// SIMATIC S7-200 project (STEP 7-Micro/WIN), CPU 224 CN REL 02.01

SYMBOL_TABLE USUARIO1
SM2              I0.0     // Sensor magnetico extendido del cilindro retenedor
SM1              I0.1     // Sensor magnetico retraido del cilindor retenedor
SM4              I0.2     // Sensor magnetico extendido del cilindro de empuje
SM3              I0.3     // Sensor magnetico retraido del cilindor de empuje
SF               I0.4     // Sensor Fotoelectrico Final
SP               I0.5     // Sensor Fotoelectrico Superior
SP1              I0.6     // Sensor Fotoelectrico Inferior
SII              I0.7     // Sensor Inductivo
SB_1             I1.2     // Pulsador de marcha
SB_2             I1.3     // Pulsador de paro
QS               I1.4     // Zeta de Emergencia
SA               I1.5     // Selector de modo
KV1              Q0.0     // Cilindro neumatico Retenedor
KV2              Q0.1     // Cilindro neumatico de empuje
HL1              Q0.7     // Señalizacion amarillo
HL2              Q1.0     // Señalizacion verde
HL3              Q1.1     // Señalizacion roja
E0               M0.0     // Estado 0
E1               M0.1     // Estado 1
E2               M0.2     // Estado 2
E3               M0.3     // Estado 3
E4               M0.4     // Estado 4
E5               M0.5     // Estado 5
EM               M0.6     // Estado de emergencia
EP               M0.7     // Estado de parada
END_SYMBOL_TABLE

ORGANIZATION_BLOCK PRINCIPAL:OB1
TITLE=COMENTARIOS DEL PROGRAMA
BEGIN
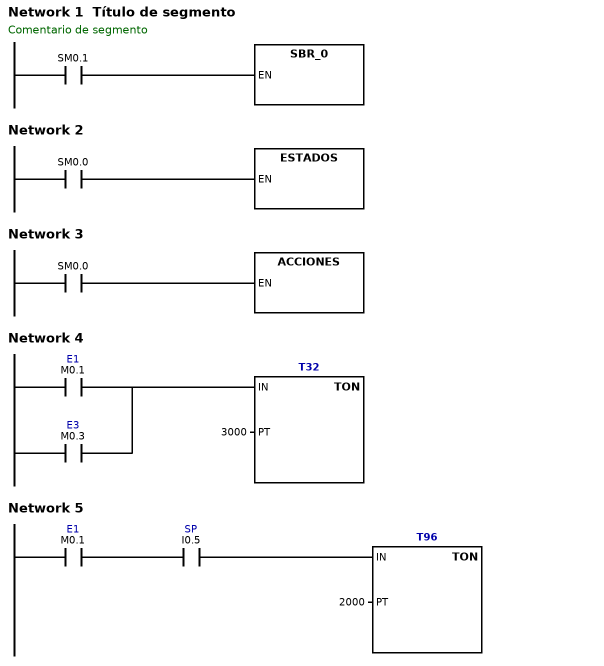
Network 1 // Título de segmento
// Comentario de segmento
LD     SM0.1
CALL   SBR_0:SBR0
Network 2
LD     SM0.0
CALL   ESTADOS:SBR1
Network 3
LD     SM0.0
CALL   ACCIONES:SBR2
Network 4
LD     E1:M0.1
O      E3:M0.3
TON    T32, 3000
Network 5
LD     E1:M0.1
A      SP:I0.5
TON    T96, 2000
END_ORGANIZATION_BLOCK

SUBROUTINE_BLOCK SBR_0:SBR0
TITLE=COMENTARIOS DE LA SUBRUTINA
BEGIN
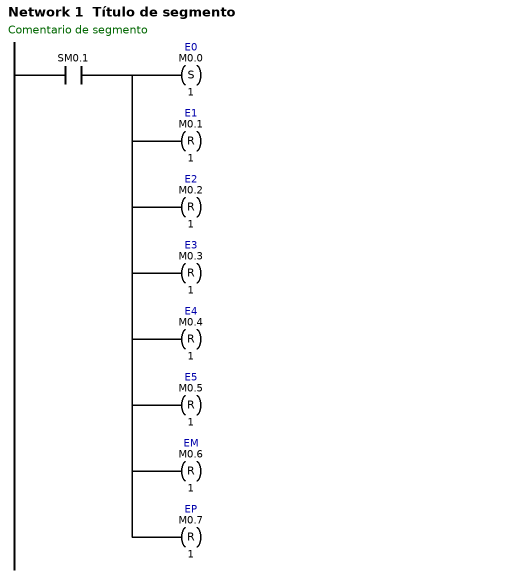
Network 1 // Título de segmento
// Comentario de segmento
LD     SM0.1
S      E0:M0.0, 1
R      E1:M0.1, 1
R      E2:M0.2, 1
R      E3:M0.3, 1
R      E4:M0.4, 1
R      E5:M0.5, 1
R      EM:M0.6, 1
R      EP:M0.7, 1
END_SUBROUTINE_BLOCK

SUBROUTINE_BLOCK ESTADOS:SBR1
TITLE=COMENTARIOS DE LA SUBRUTINA
BEGIN
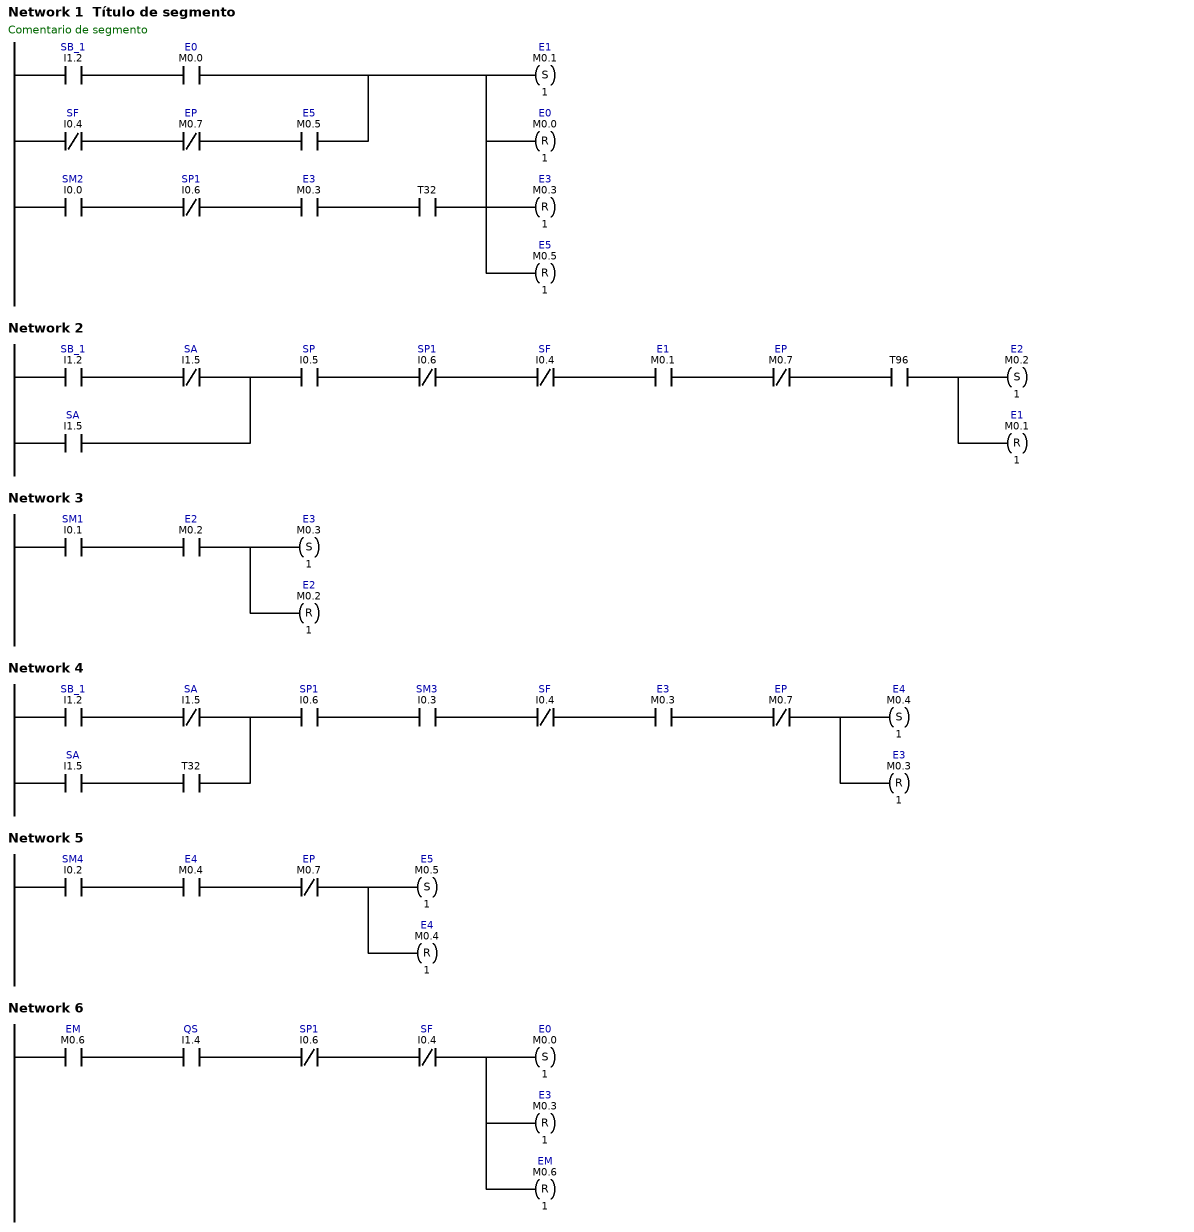
Network 1 // Título de segmento
// Comentario de segmento
LD     SB_1:I1.2
A      E0:M0.0
LDN    SF:I0.4
AN     EP:M0.7
A      E5:M0.5
OLD
LD     SM2:I0.0
AN     SP1:I0.6
A      E3:M0.3
A      T32
OLD
S      E1:M0.1, 1
R      E0:M0.0, 1
R      E3:M0.3, 1
R      E5:M0.5, 1
Network 2
// (network saved uncompiled; LAD cells follow)
// row 0: c0 -| |- SB_1:I1.2  c1 -|/|- SA:I1.5 v  c2 -| |- SP:I0.5  c3 -|/|- SP1:I0.6  c4 -|/|- SF:I0.4  c5 -| |- E1:M0.1  c6 -|/|- EP:M0.7  c7 -| |- T96 v  c8 -(S) E2:M0.2, 1
// row 1: c0 -| |- SA:I1.5  c1 -- ^  c7 ^  c8 -(R) E1:M0.1, 1
Network 3
LD     SM1:I0.1
A      E2:M0.2
S      E3:M0.3, 1
R      E2:M0.2, 1
Network 4
LD     SB_1:I1.2
AN     SA:I1.5
LD     SA:I1.5
A      T32
OLD
A      SP1:I0.6
A      SM3:I0.3
AN     SF:I0.4
A      E3:M0.3
AN     EP:M0.7
S      E4:M0.4, 1
R      E3:M0.3, 1
Network 5
LD     SM4:I0.2
A      E4:M0.4
AN     EP:M0.7
S      E5:M0.5, 1
R      E4:M0.4, 1
Network 6
LD     EM:M0.6
A      QS:I1.4
AN     SP1:I0.6
AN     SF:I0.4
S      E0:M0.0, 1
R      E3:M0.3, 1
R      EM:M0.6, 1
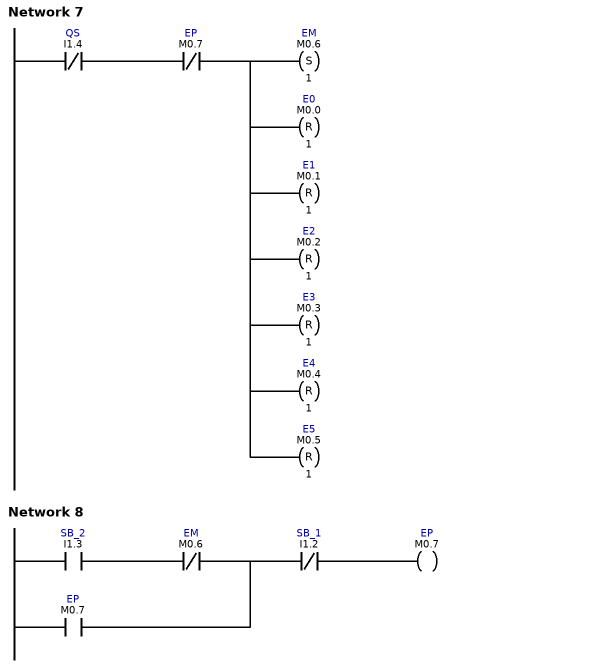
Network 7
LDN    QS:I1.4
AN     EP:M0.7
S      EM:M0.6, 1
R      E0:M0.0, 1
R      E1:M0.1, 1
R      E2:M0.2, 1
R      E3:M0.3, 1
R      E4:M0.4, 1
R      E5:M0.5, 1
Network 8
LD     SB_2:I1.3
AN     EM:M0.6
O      EP:M0.7
AN     SB_1:I1.2
=      EP:M0.7
END_SUBROUTINE_BLOCK

SUBROUTINE_BLOCK ACCIONES:SBR2
TITLE=COMENTARIOS DE LA SUBRUTINA
BEGIN
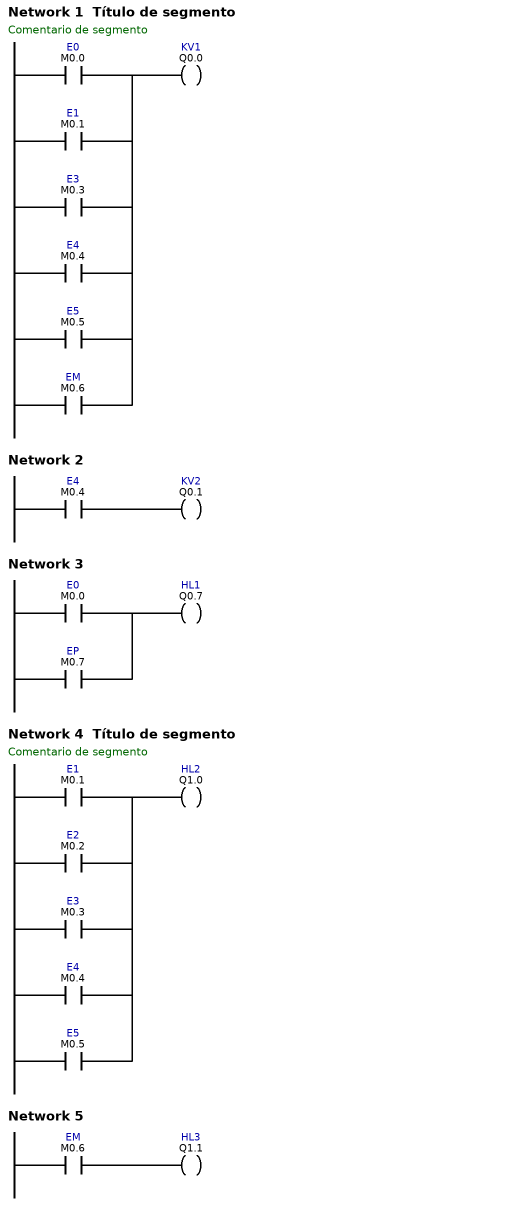
Network 1 // Título de segmento
// Comentario de segmento
LD     E0:M0.0
O      E1:M0.1
O      E3:M0.3
O      E4:M0.4
O      E5:M0.5
O      EM:M0.6
=      KV1:Q0.0
Network 2
LD     E4:M0.4
=      KV2:Q0.1
Network 3
LD     E0:M0.0
O      EP:M0.7
=      HL1:Q0.7
Network 4 // Título de segmento
// Comentario de segmento
LD     E1:M0.1
O      E2:M0.2
O      E3:M0.3
O      E4:M0.4
O      E5:M0.5
=      HL2:Q1.0
Network 5
LD     EM:M0.6
=      HL3:Q1.1
END_SUBROUTINE_BLOCK
